Fanuc KAREL source: KT00169.KL

PROGRAM KT00169
%NOLOCKGROUP
VAR
  R1: REAL
  I2: INTEGER
  OUT: INTEGER
BEGIN
  R1 = 2.0
    I2 = 3
  OUT = R1 MOD I2
END KT00169
